(* IEC 61131-3 sources: daoli-st-library/_quarantine/R84, 3 files *)

(* ---- FC_DL_FluidBedDryLossCalc.st ---- *)
(*
  DL Factory R84 | FC_DL_FluidBedDryLossCalc
  功能：算流化床干燥失重 LOD 与干基含水率，并按 2% 典型限判合格
  开源溯源：无（clean-room 自研，依据公开工艺公式，来源=行业通用公式，许可证=MIT，借鉴点=公式结构）
  规则：R1-R16 全遵守
*)
FUNCTION FC_DL_FluidBedDryLossCalc : REAL
VAR_INPUT
    fWetG : REAL := 100.0; // 干燥前湿重 [g] / wet mass before drying [g]
    fDryG : REAL := 98.0; // 干燥后干重 [g] / dry mass after drying [g]
    fLimitPct : REAL := 2.0; // LOD 合格上限（典型 2%） [%] / LOD acceptance limit [%]
END_VAR
VAR_OUTPUT
    fWaterPct : REAL; // 干基含水率（水分/干固） [%] / moisture on dry basis [%]
    xPass : BOOL; // LOD 判合格 [-] / LOD passed [-]
    xValid : BOOL; // 计算结果有效标志 [-] / calculation valid flag [-]
END_VAR
VAR
    fLossG : REAL; // 失重质量 [g] / mass loss [g]
    fLodPct : REAL; // 湿基失重中间量 [%] / wet basis loss intermediate [%]
END_VAR

// 段 1｜出口预置（R256）
FC_DL_FluidBedDryLossCalc := -1.0; // 哨兵返回 -1（无效） [-] / sentinel return -1, invalid [-]
fWaterPct := 0.0; // 含水率预置零 [%] / moisture preset zero [%]
xPass := FALSE; // 合格位预置 FALSE [-] / pass preset false [-]
xValid := FALSE; // 计算完成前不认结果 [-] / unusable before calculation [-]

// 段 2｜非有限拦截 + 质量域闸（R4/R20）
IF NOT (fWetG > -1.0E30 AND fWetG < 1.0E30) OR NOT (fDryG > -1.0E30 AND fDryG < 1.0E30) OR NOT (fLimitPct > -1.0E30 AND fLimitPct < 1.0E30) THEN
    RETURN; // 任一入参为 NaN/Inf 一律拒绝 [-] / any NaN or Inf input rejected [-]
END_IF
IF fWetG < 1.0E-9 OR fDryG < 0.0 THEN
    RETURN; // 湿重分母闸 + 干重非负闸 [g] / wet mass denominator gate and non negative dry mass [g]
END_IF
IF fDryG > fWetG THEN
    RETURN; // 干重大于湿重违反质量守恒，拒算 [g] / dry above wet violates mass balance [g]
END_IF
IF fLimitPct <= 0.0 THEN
    RETURN; // 限值正域闸 [%] / positive limit gate [%]
END_IF

// 段 3｜LOD = (湿重 − 干重) / 湿重 × 100
fLossG := fWetG - fDryG; // g − g = g / [g] minus [g] = [g]
fLodPct := (fLossG / fWetG) * 100.0; // g ÷ g × 100 = % / [g] / [g] × 100 = [%]
IF NOT (fLodPct > -1.0E30 AND fLodPct < 1.0E30) THEN
    RETURN; // 结果非有限再拦一次 [-] / second finiteness gate [-]
END_IF

// 段 4｜干基含水率 = 失重 / 干固 × 100（与湿基 LOD 区分）
IF fDryG >= 1.0E-9 THEN
    fWaterPct := (fLossG / fDryG) * 100.0; // g ÷ g × 100 = % / [g] / [g] × 100 = [%]
ELSE
    fWaterPct := -1.0; // 干重趋零：干基含水率无界，置哨兵 [%] / zero dry mass gives no finite basis [%]
END_IF
xPass := fLodPct <= fLimitPct; // 直比上限，禁浮点等值 [-] / direct compare against the limit [-]
xValid := TRUE; // 链路有效 [-] / chain valid [-]
FC_DL_FluidBedDryLossCalc := fLodPct; // 返回 LOD [%] / return the LOD [%]
END_FUNCTION

(* ---- FB_DL_ReactorHeatupProfile.st ---- *)
(*
  DL Factory R84 | FB_DL_ReactorHeatupProfile
  功能：反应釜升温程序段执行，按斜率追踪设定值并带超调抑制带与保温计时
  开源溯源：无（clean-room 自研，依据公开工艺公式，来源=行业通用公式，许可证=MIT，借鉴点=公式结构）
  规则：R1-R16 全遵守
*)
TYPE E_DL_ReactorHeatState :
(
    eIdle := 0, // 空闲待启动 [-] / idle [-]
    eRamp := 1, // 升温斜率段 [-] / heating ramp phase [-]
    eHold := 2, // 保温段 [-] / holding phase [-]
    eCool := 3, // 降温段 [-] / cooling phase [-]
    eDone := 4, // 完成相 [-] / done phase [-]
    eFault := 5 // 故障锁存相 [-] / fault latched phase [-]
) := eIdle;
END_TYPE

FUNCTION_BLOCK FB_DL_ReactorHeatupProfile
VAR_INPUT
    xStart : BOOL; // 程序段启动命令 [-] / profile start command [-]
    xReset : BOOL; // 复位命令，上升沿清故障码 [-] / reset command [-]
    rPv : REAL; // 釜内实测温度 [℃] / measured batch temperature [C]
    rTargetC : REAL := 120.0; // 升温目标温度 [℃] / heating target temperature [C]
    rCoolTargetC : REAL := 40.0; // 降温目标温度 [℃] / cooling target temperature [C]
    fRampKmin : REAL := 1.0; // 升温斜率 [K/min] / heating ramp rate [K/min]
    fCoolKmin : REAL := 0.5; // 降温斜率 [K/min] / cooling ramp rate [K/min]
    fBandK : REAL := 2.0; // 超调抑制带/到位带宽 [K] / overshoot suppression band [K]
    tHoldLimit : TIME := T#30M; // 保温时长 [s] / holding duration [s]
    tScan : TIME := T#100MS; // 扫描周期 [s] / scan period [s]
END_VAR
VAR_OUTPUT
    eState : E_DL_ReactorHeatState; // 当前程序段状态 [-] / current profile state [-]
    rSetpoint : REAL; // 当前温度设定值 [℃] / current temperature setpoint [C]
    iErrCode : INT; // 故障码 0=正常，601=组态非法，602=非法相位 [-] / error code, 601 config, 602 illegal phase [code]
    xInBand : BOOL; // 实测值落在设定带内 [-] / measured value inside the band [-]
END_VAR
VAR
    rtStart : R_TRIG; // 启动上升沿实例 [-] / start rising edge instance [-]
    rtReset : R_TRIG; // 复位上升沿实例 [-] / reset edge instance [-]
    tonHold : TON; // 保温计时器 [-] / holding timer [-]
    _eState : E_DL_ReactorHeatState := E_DL_ReactorHeatState.eIdle; // 内部相位（CASE 唯一写目标） [-] / internal phase [-]
    _iErr : INT; // 故障码内部锁存 [-] / latched error code [-]
    rSp : REAL; // 设定值内部量 [℃] / internal setpoint [C]
    fDtSec : REAL; // 扫描周期秒值 [s] / scan period in seconds [s]
    fStepK : REAL; // 本拍升/降温步长 [K] / step per scan [K]
    xCfgBad : BOOL; // 组态非法当拍标志 [-] / illegal configuration flag [-]
END_VAR

// 段 0｜边沿与定时器实例无条件周期刷新（R7）
rtStart(CLK := xStart); // 启动沿每拍必调 [-] / start edge every scan [-]
rtReset(CLK := xReset); // 复位沿每拍必调 [-] / reset edge every scan [-]
tonHold(IN := _eState = E_DL_ReactorHeatState.eHold, PT := tHoldLimit); // 保温相闸 [-] / holding phase gate [-]

// 段 1｜组态闸与扫描周期派生（斜率、带宽、周期必须正域）
fDtSec := LREAL_TO_REAL(TIME_TO_LREAL(tScan) / 1000.0); // ms ÷ 1000 = s / [ms] / 1000 = [s]
xCfgBad := NOT (fBandK > 1.0E-9) OR NOT (fRampKmin > 1.0E-9) OR NOT (fCoolKmin > 1.0E-9) OR NOT (fDtSec > 1.0E-9); // 带宽/斜率/周期正域闸（防除零） [-] / positive band, ramp and period gate [-]
xCfgBad := xCfgBad OR NOT (rTargetC > -1.0E30 AND rTargetC < 1.0E30) OR NOT (rPv > -1.0E30 AND rPv < 1.0E30); // 温度非有限闸 [-] / non finite temperature gate [-]
IF xCfgBad THEN
    _iErr := 601; // 组态非法码 [-] / illegal configuration code [-]
    _eState := E_DL_ReactorHeatState.eFault; // 锁存迁故障相 [-] / latch into the fault phase [-]
END_IF

// 段 2｜复位沿：清故障码与相位（R189）
IF rtReset.Q THEN
    _iErr := 0; // 清故障码 [-] / clear error code [-]
    _eState := E_DL_ReactorHeatState.eIdle; // 回空闲相 [-] / back to idle [-]
END_IF

// 段 3｜主状态机（合法事件优先于超时迁移，R275）
CASE _eState OF
    E_DL_ReactorHeatState.eIdle: // 空闲相：设定值初始化为实测值（无扰切换） [-] / idle [-]
        rSp := rPv; // ℃ 直取，避免起步跳变 / take the measurement to avoid a bump [C]
        IF rtStart.Q THEN
            _eState := E_DL_ReactorHeatState.eRamp; // 启动沿进升温段 [-] / start edge enters the ramp [-]
        END_IF
    E_DL_ReactorHeatState.eRamp: // 升温斜率段 [-] / heating ramp [-]
        fStepK := (fRampKmin * fDtSec) / 60.0; // K/min × s ÷ 60 = K / [K/min] × [s] / 60 = [K]
        IF (rSp + fStepK) >= rTargetC THEN
            rSp := rTargetC; // 到顶钳位，抑制超调 [-] / clamp at the target, suppress overshoot [-]
        ELSE
            rSp := rSp + fStepK; // K + K = K / [K] + [K] = [K]
        END_IF
        IF (rTargetC - rSp) < 1.0E-9 THEN
            _eState := E_DL_ReactorHeatState.eHold; // 设定值到顶转保温段 [-] / setpoint reached leads to hold [-]
        END_IF
    E_DL_ReactorHeatState.eHold: // 保温段：设定值锁定为目标 [-] / holding [-]
        rSp := rTargetC; // 锁定目标值 [℃] / lock the target [C]
        IF tonHold.Q THEN
            _eState := E_DL_ReactorHeatState.eCool; // 保温时长到转降温段 [-] / hold done leads to cooling [-]
        END_IF
    E_DL_ReactorHeatState.eCool: // 降温段 [-] / cooling [-]
        fStepK := (fCoolKmin * fDtSec) / 60.0; // K/min × s ÷ 60 = K / [K/min] × [s] / 60 = [K]
        IF (rSp - fStepK) <= rCoolTargetC THEN
            rSp := rCoolTargetC; // 到底钳位，抑制过冷 [-] / clamp at the floor, suppress undershoot [-]
        ELSE
            rSp := rSp - fStepK; // K − K = K / [K] minus [K] = [K]
        END_IF
        IF (rSp - rCoolTargetC) < 1.0E-9 THEN
            _eState := E_DL_ReactorHeatState.eDone; // 降到目标转完成相 [-] / cooled down leads to done [-]
        END_IF
    E_DL_ReactorHeatState.eDone: // 完成相 [-] / done [-]
        rSp := rCoolTargetC; // 保持终值 [℃] / hold the final value [C]
        IF NOT xStart THEN
            _eState := E_DL_ReactorHeatState.eIdle; // 命令撤销回空闲 [-] / command released returns to idle [-]
        END_IF
    E_DL_ReactorHeatState.eFault: // 故障相：码值锁存回放，仅复位沿出 [-] / fault, exit only on reset [-]
        ; // 锁存回放（R28） [-] / replay the latch only [-]
ELSE
    _iErr := 602; _eState := E_DL_ReactorHeatState.eFault; // 非法相位兜底 [-] / illegal phase fallback [-]
END_CASE

// 段 4｜出口映射（名实双出口，同源赋值）
eState := _eState; // 状态出口 [-] / state outlet [-]
rSetpoint := rSp; // 设定值出口 [℃] / setpoint outlet [C]
iErrCode := _iErr; // 故障码出口（锁存值） [-] / error code outlet [-]
xInBand := (ABS(rPv - rSp) <= fBandK) AND NOT xCfgBad; // K 差值与带宽直比，组态非法时强制 FALSE（连续量出口防护） [-] / band compare with a config fault override [-]
END_FUNCTION_BLOCK

(* ---- FB_DL_ToolMagazinePosSeq.st ---- *)
(*
  DL Factory R84 | FB_DL_ToolMagazinePosSeq
  功能：刀库就近寻刀定位时序，含双向索引差取小择向与旋转/锁紧双超时
  开源溯源：无（clean-room 自研，依据公开工艺公式，来源=行业通用公式，许可证=MIT，借鉴点=公式结构）
  规则：R1-R16 全遵守
*)
TYPE E_DL_TmagState :
(
    eIdle := 0, // 空闲待命 [-] / idle [-]
    eSearch := 1, // 就近择向计算相 [-] / nearest slot evaluation phase [-]
    eRotate := 2, // 刀盘旋转相 [-] / magazine rotation phase [-]
    eLockCheck := 3, // 锁紧确认相 [-] / lock confirmation phase [-]
    eReady := 4, // 定位完成相 [-] / positioned phase [-]
    eFault := 5 // 故障锁存相 [-] / fault latched phase [-]
) := eIdle;
END_TYPE

FUNCTION_BLOCK FB_DL_ToolMagazinePosSeq
VAR_INPUT
    xStart : BOOL; // 寻刀启动命令 [-] / seek start command [-]
    xReset : BOOL; // 复位命令（上升沿清故障码） [-] / reset command [-]
    iReqSlot : INT; // 请求刀位序号（0 基） [个] / requested slot index, zero based [count]
    iCurSlot : INT; // 当前刀位序号（0 基） [个] / current slot index, zero based [count]
    iSlotCnt : INT; // 刀库总刀位数（1~200） [个] / total slot count [count]
    xRotInPos : BOOL; // 旋转到位反馈 [-] / rotation in position feedback [-]
    xLocked : BOOL; // 刀盘锁紧确认 [-] / magazine locked confirmation [-]
    tRotLimit : TIME := T#20S; // 旋转到位超时门限 [s] / rotation timeout [s]
    tLockLimit : TIME := T#3S; // 锁紧确认超时门限 [s] / lock timeout [s]
END_VAR
VAR_OUTPUT
    eState : E_DL_TmagState; // 当前时序状态 [-] / current sequence state [-]
    iTargetSlot : INT; // 择定的目标刀位序号（0 基） [个] / resolved target slot [count]
    iErrCode : INT; // 故障码 0=正常，301~304 [-] / error code, 301 to 304 [code]
    xReady : BOOL; // 定位完成（可换刀） [-] / positioned and ready [-]
    iDirCtrl : INT; // 择向指令出口 1=正转 −1=反转 0=未定 [-] / direction command outlet, 1 forward -1 reverse 0 undecided (R583)
END_VAR
VAR
    rtStart : R_TRIG; // 启动上升沿实例 [-] / start rising edge instance [-]
    rtReset : R_TRIG; // 复位上升沿实例 [-] / reset rising edge instance [-]
    tonRot : TON; // 旋转到位超时定时器 [-] / rotation timeout timer [-]
    tonLock : TON; // 锁紧确认超时定时器 [-] / lock timeout timer [-]
    _eState : E_DL_TmagState := E_DL_TmagState.eIdle; // 内部相位（CASE 唯一写目标） [-] / internal phase [-]
    _iErr : INT; // 故障码内部锁存 [-] / latched error code [-]
    iDiff : INT; // 正向索引差（已取绝对值） [个] / forward absolute index difference [count]
    iAlt : INT; // 反向索引差 [个] / reverse index difference [count]
    iDir : INT; // 择向结果 1=正转 −1=反转 [-] / chosen direction [-]
END_VAR

// 段 0｜边沿与定时器实例无条件周期刷新（R7）
rtStart(CLK := xStart); // 启动沿每拍必调 [-] / start edge called every scan [-]
rtReset(CLK := xReset); // 复位沿每拍必调 [-] / reset edge called every scan [-]
tonRot(IN := _eState = E_DL_TmagState.eRotate, PT := tRotLimit); // 旋转相闸 + 无条件调用 [-] / rotation timer, unconditional [-]
tonLock(IN := _eState = E_DL_TmagState.eLockCheck, PT := tLockLimit); // 锁紧相闸 + 无条件调用 [-] / lock timer, unconditional [-]

// 段 0｜出口预置（R256）：择向指令每拍先归未定，由 eSearch 单点重赋
iDir := 0; // 未择向 [-] / undecided direction [-]

// 段 1｜复位沿：清故障码与相位（保持量不含 Prev/Acc/Latch，R189）
IF rtReset.Q THEN
    _iErr := 0; // 清故障码 [-] / clear error code [-]
    _eState := E_DL_TmagState.eIdle; // 回空闲相 [-] / back to idle [-]
END_IF

// 段 2｜主状态机（合法事件优先于超时迁移，R275）
CASE _eState OF
    E_DL_TmagState.eIdle: // 空闲相 [-] / idle [-]
        IF rtStart.Q THEN
            _eState := E_DL_TmagState.eSearch; // 启动沿进择向相 [-] / start edge enters evaluation [-]
        END_IF
    E_DL_TmagState.eSearch: // 就近择向：两方向索引差取小（有符号差显式取模，R271 禁单侧 ABS） [-] / nearest direction [-]
        IF (iSlotCnt < 1) OR (iSlotCnt > 200) OR (iReqSlot < 0) OR (iReqSlot >= iSlotCnt) OR (iCurSlot < 0) OR (iCurSlot >= iSlotCnt) THEN
            _iErr := 301; _eState := E_DL_TmagState.eFault; // 刀位组态越界 [-] / slot index out of range [-]
        ELSE
            iDiff := iReqSlot - iCurSlot; // 有符号差先求再取模 [个] / signed difference [count]
            IF iDiff < 0 THEN
                iDiff := -iDiff; // 双侧直比：负数显式取反 [个] / take the magnitude explicitly [count]
            END_IF
            iAlt := iSlotCnt - iDiff; // 反向圈数 = 总数 − 正向步数 [个] / reverse count [count]
            IF iDiff <= iAlt THEN
                iDir := 1; // 正向不多于反向，取正转 [-] / forward is not longer [-]
            ELSE
                iDir := -1; // 反向更短，取反转 [-] / reverse is shorter [-]
            END_IF
            iTargetSlot := iReqSlot; // 输出择定目标刀位 [个] / export the resolved slot [count]
            _eState := E_DL_TmagState.eRotate; // 择向完成立即转旋转相 [-] / evaluation leads to rotation [-]
        END_IF
    E_DL_TmagState.eRotate: // 旋转相（iDir 供执行层决定正/反转） [-] / rotation [-]
        IF xRotInPos AND NOT tonRot.Q THEN
            _eState := E_DL_TmagState.eLockCheck; // 到位转锁紧确认 [-] / in position leads to lock check [-]
        ELSIF tonRot.Q THEN
            _iErr := 302; _eState := E_DL_TmagState.eFault; // 旋转到位超时 [-] / rotation timeout [-]
        END_IF
    E_DL_TmagState.eLockCheck: // 锁紧确认相（上锁类安全相，入相复检无故障） [-] / lock check [-]
        IF xLocked AND NOT tonLock.Q THEN
            _eState := E_DL_TmagState.eReady; // 锁紧确认转完成相 [-] / locked leads to ready [-]
        ELSIF tonLock.Q THEN
            _iErr := 303; _eState := E_DL_TmagState.eFault; // 锁紧确认超时 [-] / lock timeout [-]
        END_IF
    E_DL_TmagState.eReady: // 定位完成相：保持刀位，命令撤销即回空闲 [-] / ready [-]
        IF NOT xStart THEN
            _eState := E_DL_TmagState.eIdle; // 命令撤销回空闲 [-] / command released returns to idle [-]
        END_IF
    E_DL_TmagState.eFault: // 故障相：码值锁存回放，仅复位沿出 [-] / fault, exit only on reset [-]
        ; // 锁存回放（读己不改值，R28） [-] / replay the latch only, no re-inference [-]
ELSE
    _iErr := 304; _eState := E_DL_TmagState.eFault; // 非法相位兜底 [-] / illegal phase fallback [-]
END_CASE

// 段 3｜出口映射（名实双出口，同源赋值）
eState := _eState; // 状态出口 [-] / state outlet [-]
iErrCode := _iErr; // 故障码出口（锁存值） [-] / error code outlet [-]
iDirCtrl := iDir; // 择向结果出口（原先仅内部量，R583 补出口） [-] / direction outlet, previously internal only [-]
xReady := _eState = E_DL_TmagState.eReady; // 完成位 = 完成相镜像 [-] / ready mirrors the ready phase [-]
END_FUNCTION_BLOCK
